Staubli VAL3: deleteProgItem.pgx

public program deleteProgItem(string x_sKey, string x_sItem, bool& x_bToSave)
  local bool l_bResult
  local bool l_bResult1
  local num l_nIndex
begin
  if x_sItem!=""
    l_bResult=userPageConfirm("是否删除"+x_sItem+"?")
    if l_bResult
      toNum(x_sItem,l_nIndex,l_bResult1)
      if l_nIndex==0 and size(progTemp:pProgItem[x_sKey].pProgTemplate)<2
        userPageAlert("数组元素数量需大于0")
      else
        delete(progTemp:pProgItem[x_sKey].pProgTemplate[l_nIndex])
        //progTemp:libSave()
        x_bToSave=true
      endIf
    endIf
  else
    userPageAlert("未选中有效项目!")
  endIf
end
